Fanuc KAREL source: KT00132.KL

PROGRAM KT00132
%NOLOCKGROUP
VAR
  I1: INTEGER
  R2: REAL
  OUT: REAL
BEGIN
  I1 = 2
    R2 = 3.0
  OUT = I1 DIV R2
END KT00132
